// TIA Portal V21 export
DATA_BLOCK "SafetyData"   // DB3, F_DB
{ S7_Optimized_Access := 'TRUE' }
// Fail-safe data shared by the safety program and read by the standard program.
   VAR
      released : Bool;
      limit : Int := 12;
   END_VAR
BEGIN
END_DATA_BLOCK
